(* IEC 61131-3 sources: Test-Git_ESME26/TestProgettoESME_26.fbsproj/PacDriveLib Migration/Motion/Control/Brake/FB_BrakeReleaseSet.fb.st^, 3 files *)

(* ---- ifBrake.prop.st ---- *)
PROPERTY ifBrake : DDI.IF_Brake
__SETTERDECLARATION__
VAR
END_VAR
__SETTERIMPLEMENTATION__
ifBrake_loc := ifBrake;

(* ---- xDone.prop.st ---- *)
PROPERTY xDone : BOOL
__GETTERDECLARATION__
VAR
END_VAR
__GETTERIMPLEMENTATION__
xDone := xDone_loc;
__SETTERDECLARATION__
VAR
END_VAR
__SETTERIMPLEMENTATION__
xDone_loc := xDone;

(* ---- xRelease.prop.st ---- *)
PROPERTY PUBLIC xRelease : BOOL
__SETTERDECLARATION__
VAR
END_VAR
__SETTERIMPLEMENTATION__
xRelease_loc := xRelease;
